// TIA Portal V21 export
// export: Created 2026-11-21T13:31:41.2452098Z, ExportSetting WithDefaults, DisplayName Totally Integrated Automation Portal, DisplayVersion V21, DisplayName STEP 7 Professional, DisplayVersion V21, DisplayName STEP 7 Safety, DisplayVersion V21, DisplayName Tech WebApplication, DisplayVersion V21, DisplayName WinCC Basic/Comfort/Advanced, DisplayVersion V21, DisplayName WinCC Unified, DisplayVersion V21
FUNCTION_BLOCK "ClassicLad"   // FB10, LAD
TITLE = ClassicLad
VERSION : 0.1
// Ladder on a classic CPU, with global tags.
// stored: AutoNumber true, IsIECCheckEnabled false, UDAEnableTagReadback false
   VAR_INPUT
      enable : Bool;
   END_VAR
   VAR_OUTPUT
      running : Bool;
   END_VAR
   VAR DB_SPECIFIC
      latched : Bool;
   END_VAR
BEGIN

REGION Network 1: Run the motor
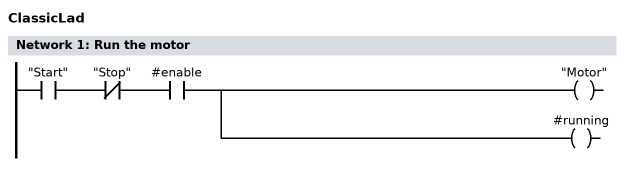
   RUNG wire#powerrail
      Contact( "Start" )
      I_Contact( "Stop" )
      Contact( #enable )
      wire#w1
      Coil( "Motor" )
   END_RUNG
   RUNG wire#w1
      Coil( #running )
   END_RUNG
   // the same network as SCL:
   "Motor" := "Start" AND NOT "Stop" AND #enable;
   #running := "Motor";
END_REGION
END_FUNCTION_BLOCK
